Fanuc KAREL source: KA00205.KL

PROGRAM KA00205
%NOLOCKGROUP
VAR
  SRC: ARRAY[4] OF VECTOR
  DST: ARRAY[4] OF VECTOR
BEGIN
  DST = SRC
END KA00205
